(* IEC 61131-3 sources: s7-to-codesys/src/POUs/S7Compat/F_S5CountDown, 2 files *)

(* ---- F_S5CountDown.decl.st ---- *)
// Назначение: CD C n — счёт вниз счётчика S5: по фронту RLO 0 → 1 значение −1, не меньше 0 (AWL_e.pdf,
//             гл. 4). Возвращает значение после инструкции.
// Автор:      kr0nsch
// Версия:     1.2.0
// Документ:   docs/MAPPING_STL.md, правило s5.counter
FUNCTION F_S5CountDown : INT
VAR_IN_OUT
    stCounter : ST_S5Counter;   // счётчик (GVL_S5Counters.aCounter[n])
END_VAR
VAR_INPUT
    xRlo : BOOL;                // RLO перед инструкцией
END_VAR

(* ---- F_S5CountDown.impl.st ---- *)
IF xRlo AND NOT stCounter.xRloDown AND stCounter.iValue > 0 THEN
    stCounter.iValue := stCounter.iValue - 1;
END_IF
stCounter.xRloDown := xRlo;
F_S5CountDown := stCounter.iValue;
